(* Logix 5000 project; controller R400_500_XLS vendor 1 type 14 code 216 rev 31.11; software revision 31.01; part 2 of 32 *)

PROGRAM MainProgram   (* main routine MainRoutine *)
VAR
   Abort1 : DINT := 1;   // Not Used
        .0   // Initial step
        .1   // Remove stop condition
        .10   // Call module to fill sump Close Rcvry Tank Drain Valve
        .12   // Drain Rcvry Tank
        .14   // Call FC13 Drain Sump
        .16   // Sump draining phase is process
        .18   // Abort Completed Display Ready Mode screen
        .2   // No Recovery Tank Option or Recoverytank option and treament is Drying or Venting Reset Functions prior to drain sump
        .21   // Reset Functions
        .22   // Reset Functions prior to drain Rcvry Tank
        .24   // Reset Functions prior to drain sump
        .26   // Reset Functions prior to drain Rcvry Tank
        .28   // Reset Functions prior to drain sump
        .31   // Start Abort Sequence
        .4   // Check Filling Port
        .6   // Reset Functions prior to drain Rcvry Tank
        .8   // Reset Functions prior to fill sump
   Abort2 : SINT := 33;
        .0   // Initial Step
        .1   // Drying or Venting treatment is running Reset Functions prior to Vent Chamber
        .2   // Drying or Venting Treat. was running Exhaust Chamber (Abort Sequence) Enrg. Fan
        .5   // Initial Step
        .6   // Recirc. or F. Rinse Treat. was running Exhaust Chamber (Abort Sequence)
   Alarm : SINT := 1;   // Wait 3 seconds
        .0   // Initial step. No alarm detected.
        .1   // Alarm detected. Stop the cycle
        .2   // The alarm is acknowledged
        .3   // Display RESUME button
        .5   // Transition
        .6   // Transition
        .7   // Run mode
   AlarmAcked : BOOL;   // Alarm has been acked
   AlarmFlag : DINT;   // Active alarm flag
        .1   // Load door did not open flag
        .10   // Pure water tank safety water level reached
        .11   // Sump too long to fill
        .12   // Sump drain too long
        .13   // Sump too long to heat
        .14   // Sump RTD defective
        .15   // Sump temperature too high
        .16   // Pure water tank too long to fill
        .17   // Pure water tank drain too long
        .18   // Pure Water Tank too long to heat
        .19   // Pure Water Tank RTD defective
        .2   // Load door did not close flag
        .20   // Pure water tank temperature too high
        .21   // Pure water tank failed to dump
        .22   // Chemical Container 1 empty
        .23   // Chemical Container 2 empty
        .24   // Chemical Container 3 empty
        .25   // Chemical Container 4 empty
        .26   // Drying temperature not reached
        .27   // Chemical injection conductivity setpoint not reached
        .28   // Final rinse conductivity setpoint not reached
        .29   // Final rinse conductivity system defective
        .3   // Load door obstructed
        .30   // Chemcial conductivity system defective
        .31   // Pressure Transmitter defective
        .4   // Load door open
        .5   // Unload door did not open
        .6   // Unload door did not close
        .7   // Unload Door Obstructed
        .8   // Unload door Open
        .9   // Sump safety level reached
   AlarmFlag1 : DINT;
        .0   // Pump pressure too low
        .1   // Motor overload detected
        .10   // Waiting For Pure Water Filling Authorization
        .11   // Audit Trail Low Storage Memory
        .2   // Maintenance due
        .3   // Both doors open
        .4   // Drying RTD defective
        .5   // Master control relay deactivated
        .6   // PURE WATER TANK TEMPERATURE ABOVE TEMPERATURE RANGE ALLOWED
        .7   // PURE WATER TANK TEMPERATURE UNDER TEMPERATURE RANGE ALLOWED
        .8   // BATTERY LOW
        .9   // I/O Communication has been lost
   AlarmMuted : BOOL;
   AlarmTran0 : BOOL;   // Transition from step 3 to step 0
   Ashutdown : SINT := 1;   // Not Used
        .0   // Initial Step
        .1   // Call manual shutdown function Start signal from the automatic shutdown requirement
        .2   // Wait activation of Wake button (initial step of OPR-13)
        .3   // Enabled door printout and wait opening of the door
        .4   // Door is open
        .5   // Unloading completed
        .6   // Accept/Reject Cycle
   bAlrm : BOOL[64];
        [10]   // PURE WATER TANK TOO LONG TO DRAIN (trigger)
        [11]   // SUMP TOO LONG TO FILL (trigger)
        [12]   // SUMP TOO LONG TO HEAT (trigger)
        [13]   // SUMP DRAIN TOO LONG (trigger)
        [14]   // Chemical container 1 low
        [15]   // Chemical container 2 low
        [16]   // Chemical container 3 low
        [17]   // Chemical container 4 low
        [18]   // ALARM PURE WATER TANK TOO LONG TO FILL (trigger)
        [19]   // Pure water tank too long to heat
        [1]   // ALARM LOAD DOOR OBSTRUCTED (trigger)
        [20]   // ALARM PURE WATER TANK FAIL TO DUMP (trigger)
        [21]   // PURE WATER TANK TOO LONG TO DRAIN
        [22]   // Drying temperature not reached (trigger)
        [23]   // Chemical container 1 low
        [24]   // Chemical container 2 low
        [25]   // Chemical container 3 low
        [26]   // Chemical container 4 low
        [27]   // Conductivity is too long to reach set point
        [28]   // Final Rinse cond. sp not reached
        [29]   // Chemical container 1 low
        [2]   // ALARM LOAD DOOR DID NOT OPEN (trigger)
        [30]   // Chemical container 2 low
        [31]   // Chemical container 3 low
        [32]   // Chemical container 4 low
        [3]   // ALARM LOAD DOOR DID NOT CLOSE (trigger)
        [4]   // Reserved Load door open
        [5]   // ALARM UNLOAD DOOR OBSTRUCTED (trigger)
        [6]   // ALARM UNLOAD DOOR DID NOT OPEN (trigger)
        [7]   // ALARM UNLOAD DOOR DID NOT CLOSE (trigger)
        [8]   // Reserved Unload Door Open
        [9]   // SUMP TOO LONG TO DRAIN (trigger)
   bChangeFromNonHeatedToHeated : BOOL;
   bResetAllCycle : BOOL;
   bResetServiceMode : BOOL;
   CalCond : SINT;
        .1   // Calibration Enabled bit
        .2   // Wait for low calibration value
        .3   // Set Low value and Wait for High value
        .4   // Set High value and Verify Calibration
   CalFrinseCond : SINT;
        .1   // Calibration Enable bit
        .2   // Wait for low calibration value
        .3   // Set Low value and Wait for High value
        .4   // Set High value and Verify Calibration
   Calib : SINT;
        .0   // Enter Low Value
        .1   // Enter High Value
        .2   // Verify Calibration
   CalibCnt : SINT := 2;   // Calibration Step Counter
   CalibCondCnt : SINT;
   CalibData : UDT_SCALE[8] := ([0].InputMin := 213, [0].InputMax := 1207, [0].ScaledMin := 218.0, [0].ScaledMax := 1212.0, [0].DfInputMax := 1000, [0].DfScaledMax := 1000, [0].Input := 212, [0].Output := 21.7, [1].InputMin := 234, [1].InputMax := 1204, [1].ScaledMin := 239.0, [1].ScaledMax := 1210.0, [1].DfInputMax := 1000, [1].DfScaledMax := 1000, [1].Input := 222, [1].Output := 22.698767, [2].InputMin := 223, [2].InputMax := 1205, [2].ScaledMin := 228.0, [2].ScaledMax := 1210.0, [2].DfInputMax := 1000, [2].DfScaledMax := 1000, [2].Input := 214, [2].Output := 21.9, [3].InputMin := 4000, [3].InputMax := 20000, [3].ScaledMax := 60.0, [3].DfInputMin := 4000, [3].DfInputMax := 20000, [3].DfScaledMax := 60, [3].Input := 12566, [3].Output := 32.122498, [4].InputMin := 4000, [4].InputMax := 20000, [4].ScaledMax := 100.0, [4].DfInputMin := 4000, [4].DfInputMax := 20000, [4].DfScaledMax := 100, [4].Input := 9495, [4].Output := 34.34375, [5].InputMin := 4000, [5].InputMax := 20000, [5].ScaledMax := 100.0, [5].DfInputMin := 4000, [5].DfInputMax := 20000, [5].DfScaledMax := 100, [5].Input := 4000, [7].InputMin := 223, [7].InputMax := 1205, [7].ScaledMin := 228.0, [7].ScaledMax := 1210.0, [7].DfInputMax := 1000, [7].DfScaledMax := 1000, [7].Input := 302, [7].Output := 30.7);
        [0]   // Sump RTD Calibration data
        [1]   // Dry RTD Calibration data
        [2]   // PWT RTD Calibration data
        [3]   // Pressure Calibration data
        [4]   // Final Rinse Channel calibration data
        [5]   // Chemical Channe calibration data
        [6]   // Spare channel
        [7]   // Reserved for printouts
   CalibEnabled : BOOL;   // RTD Calibration Enabled bit
   CalibFrinseCondCnt : SINT;
   CalibIndex : DINT := 1;   // Calibration Pointer
   CalibPressCnt : SINT := 2;
   CalPressure : SINT;
   Change_PrintPtr_Value : BOOL;
   Chem_Pump : UDT_CHEM_PUMP[4] := ([0].FlowRate := 270, [1].FlowRate := 270, [2].FlowRate := 270, [3].FlowRate := 270);   // Chemical Pump flow rate
        [0].FlowRate   // Flow rate of Pump 1
        [1].FlowRate   // Flow rate of Pump 2
        [2].FlowRate   // Flow rate of Pump 3
        [3].FlowRate   // Flow rate of Pump 4
   CHEMICAL_COND_MAX_TIME : DINT := 360000;   // Timeout for the conductivity based chemical injection
   CHEMICAL_PUMP_OFF_TIME : DINT[4] := ([0] := 8, [1] := 8, [2] := 8, [3] := 8);
   CHEMICAL_PUMP_ON_TIME : DINT[4] := ([0] := 2, [1] := 2, [2] := 2, [3] := 2);
   ChemPumpIndex : DINT := 1;
   ChPumpRunningTime : REAL := 42.043003;
   ClearIndex : DINT := 300;
   Condenser : INT := 1025;
        .0   // Initial step. Condenser stopped
        .1   // Condenser operating
        .10   // Initial step. Condenser stopped
        .11   // Condenser operating
   CondenserHighFlow_1 : BOOL;   // Enables the condenser high flow valve
   CondenserHighFlow_2 : BOOL;   // Enables the condenser high flow valve
   CondenserLowFlow_1 : BOOL;   // Enables the condenser low flow valve
   CondenserLowFlow_2 : BOOL;   // Enables the condenser low flow valve
   CondenserTran : INT;
        .0   // From step 0 to 1
        .1   // From step 1 to 0
        .10   // From step 10 to step 11
        .11   // From step 11 to step 10
   Critical_Alarm : BOOL;
   CURRENT_CYCLE : DINT := 11;
   CustomCycleIterator : DINT := 11;
   CycExcBuffer : UDT_CYCLE := (PW[0].Wprt := 2, PW[0].Tmin := 1, PW[1].Wprt := 2, PW[2].Wprt := 2, PW[3].Wprt := 2, WSH[0].Wprt := 2, WSH[1].Wprt := 2, WSH[2].Wprt := 2, WSH[3].Wprt := 2, WSH[4].Wprt := 2, RINSE[0].Wprt := 2, RINSE[1].Wprt := 2, RINSE[2].Wprt := 2, RINSE[3].Wprt := 2, FRINSE.Tsec := 10, FRINSE.Drn := 1, DRY.HeatSensitive := 1, Lock := 1);
   CycleDryingStandard : UDT_DRY := (Mode := 1, Tmin := 15, HiLowTemp := 1);
   CycleModifBuffer : UDT_CYCLE := (PW[0].Wprt := 2, PW[0].Tmin := 1, PW[1].Wprt := 2, PW[2].Wprt := 2, PW[3].Wprt := 2, WSH[0].Wprt := 2, WSH[1].Wprt := 2, WSH[2].Wprt := 2, WSH[3].Wprt := 2, WSH[4].Wprt := 2, RINSE[0].Wprt := 2, RINSE[1].Wprt := 2, RINSE[2].Wprt := 2, RINSE[3].Wprt := 2, FRINSE.Tsec := 10, FRINSE.Drn := 1, DRY.HeatSensitive := 1, Lock := 1);
   CycleNotEmpty : SINT;
   Cycles : UDT_CYCLE[11] := ([0].PW[0].TrtNo := 1, [0].PW[0].Wprt := 1, [0].PW[0].Tmin := 2, [0].PW[1].Wprt := 2, [0].PW[2].Wprt := 2, [0].PW[3].Wprt := 2, [0].WSH[0].Wprt := 2, [0].WSH[0].Heat := 1, [0].WSH[0].Tmp := 65.6, [0].WSH[0].Tmin := 10, [0].WSH[0].ChemUsed_1 := 1, [0].WSH[0].ChemVol_1 := 4.0, [0].WSH[1].Wprt := 2, [0].WSH[2].Wprt := 2, [0].WSH[2].Heat := 1, [0].WSH[2].Tmp := 65.6, [0].WSH[2].Tmin := 1, [0].WSH[2].ChemUsed_1 := 2, [0].WSH[2].ChemVol_1 := 4.0, [0].WSH[3].Wprt := 2, [0].WSH[4].Wprt := 2, [0].RINSE[0].Wprt := 2, [0].RINSE[0].Tmin := 4, [0].RINSE[1].Wprt := 2, [0].RINSE[1].Tmin := 8, [0].RINSE[2].Wprt := 2, [0].RINSE[3].Wprt := 2, [0].FRINSE.Heat := 1, [0].FRINSE.Tmp := 50.0, [0].FRINSE.Tsec := 10, [0].FRINSE.Nb := 1, [0].FRINSE.Recirc := 1, [0].FRINSE.Drn := 1, [0].DRY.Mode := 1, [0].DRY.Tmin := 25, [0].DRY.HiLowTemp := 1, [0].Lock := 1, [1].PW[0].Wprt := 1, [1].PW[0].Tmin := 2, [1].PW[1].Wprt := 2, [1].PW[2].Wprt := 2, [1].PW[3].Wprt := 2, [1].WSH[0].Wprt := 2, [1].WSH[0].Heat := 1, [1].WSH[0].Tmp := 65.6, [1].WSH[0].Tmin := 10, [1].WSH[0].ChemUsed_1 := 1, [1].WSH[0].ChemVol_1 := 3.90625, [1].WSH[1].Wprt := 2, [1].WSH[2].Wprt := 2, [1].WSH[3].Wprt := 2, [1].WSH[4].Wprt := 2, [1].RINSE[0].Wprt := 2, [1].RINSE[0].Tmin := 4, [1].RINSE[1].Wprt := 2, [1].RINSE[1].Heat := 1, [1].RINSE[1].Tmp := 65.6, [1].RINSE[1].Tmin := 8, [1].RINSE[2].Wprt := 2, [1].RINSE[3].Wprt := 2,
        [1].FRINSE.Heat := 1, [1].FRINSE.Tmp := 65.6, [1].FRINSE.Tsec := 10, [1].FRINSE.Nb := 2, [1].FRINSE.Drn := 1, [1].DRY.HeatSensitive := 1, [1].Lock := 1, [2].PW[0].Wprt := 2, [2].PW[0].Tmin := 2, [2].PW[1].Wprt := 2, [2].PW[2].Wprt := 2, [2].PW[3].Wprt := 2, [2].WSH[0].Wprt := 2, [2].WSH[0].Heat := 1, [2].WSH[0].Tmp := 65.6, [2].WSH[0].Tmin := 10, [2].WSH[1].Wprt := 2, [2].WSH[2].Wprt := 2, [2].WSH[3].Wprt := 2, [2].WSH[4].Wprt := 2, [2].RINSE[0].Wprt := 2, [2].RINSE[0].Tmin := 4, [2].RINSE[1].Wprt := 1, [2].RINSE[1].Tmin := 8, [2].RINSE[2].Wprt := 2, [2].RINSE[3].Wprt := 2, [2].FRINSE.Tsec := 10, [2].FRINSE.Nb := 2, [2].FRINSE.Drn := 1, [2].DRY.Mode := 1, [2].Lock := 1, [3].PW[0].Wprt := 1, [3].PW[1].Wprt := 2, [3].PW[2].Wprt := 2, [3].PW[3].Wprt := 2, [3].WSH[0].Wprt := 2, [3].WSH[0].Heat := 1, [3].WSH[0].Tmp := 65.6, [3].WSH[0].ChemUsed_1 := 1, [3].WSH[0].ChemVol_1 := 0.9765625, [3].WSH[1].Wprt := 2, [3].WSH[2].Wprt := 2, [3].WSH[3].Wprt := 2, [3].WSH[4].Wprt := 2, [3].RINSE[0].Wprt := 2, [3].RINSE[1].Wprt := 2, [3].RINSE[2].Wprt := 2, [3].RINSE[3].Wprt := 2, [3].FRINSE.Heat := 1, [3].FRINSE.Tmp := 50.0, [3].FRINSE.Tsec := 30, [3].FRINSE.Recirc := 1, [3].FRINSE.Drn := 1, [3].DRY.Mode := 1, [3].DRY.Tmin := 25, [3].DRY.HiLowTemp := 1, [3].Lock := 1, [4].PW[0].Wprt := 2, [4].PW[0].Tmin := 2, [4].PW[0].Tsec := 30,
        [4].PW[1].Wprt := 1, [4].PW[1].Tmin := 1, [4].PW[2].Wprt := 2, [4].PW[3].Wprt := 2, [4].WSH[0].Wprt := 2, [4].WSH[0].Tmin := 10, [4].WSH[0].ChemUsed_1 := 1, [4].WSH[0].ChemVol_1 := 1.953125, [4].WSH[1].Wprt := 2, [4].WSH[1].Heat := 1, [4].WSH[1].Tmp := 65.6, [4].WSH[1].Tmin := 4, [4].WSH[2].Wprt := 2, [4].WSH[2].Tmin := 10, [4].WSH[2].ChemUsed_1 := 1, [4].WSH[2].ChemVol_1 := 3.90625, [4].WSH[3].Wprt := 2, [4].WSH[4].Wprt := 2, [4].RINSE[0].Wprt := 2, [4].RINSE[1].Wprt := 2, [4].RINSE[2].Wprt := 2, [4].RINSE[3].Wprt := 2, [4].FRINSE.Heat := 1, [4].FRINSE.Tmp := 50.0, [4].FRINSE.Tsec := 30, [4].FRINSE.Recirc := 1, [4].FRINSE.Drn := 1, [4].DRY.Mode := 1, [4].Lock := 1, [5].PW[0].Wprt := 2, [5].PW[1].Wprt := 2, [5].PW[2].Wprt := 2, [5].PW[3].Wprt := 2, [5].WSH[0].Wprt := 2, [5].WSH[0].Heat := 1, [5].WSH[0].Tmp := 65.6, [5].WSH[0].ChemUsed_1 := 2, [5].WSH[0].ChemVol_1 := 16.0, [5].WSH[1].Wprt := 2, [5].WSH[2].Wprt := 2, [5].WSH[3].Wprt := 2, [5].WSH[4].Wprt := 2, [5].RINSE[0].Wprt := 2, [5].RINSE[0].Tmin := 10, [5].RINSE[1].Wprt := 2, [5].RINSE[1].Tmin := 10, [5].RINSE[2].Wprt := 2, [5].RINSE[2].Tmin := 10, [5].RINSE[3].Wprt := 2, [5].FRINSE.Heat := 1, [5].FRINSE.Tmp := 50.0, [5].FRINSE.Tsec := 30, [5].FRINSE.Recirc := 1, [5].FRINSE.Drn := 1, [5].DRY.Mode := 1, [5].DRY.Tmin := 15, [5].DRY.HiLowTemp := 1, [5].Lock := 1, [6].PW[0].Wprt := 2, [6].PW[0].Tmin := 1,
        [6].PW[1].Wprt := 2, [6].PW[2].Wprt := 2, [6].PW[3].Wprt := 2, [6].WSH[0].Wprt := 2, [6].WSH[0].Heat := 1, [6].WSH[0].Tmp := 70.0, [6].WSH[0].ChemUsed_1 := 1, [6].WSH[0].ChemVol_1 := 1.953125, [6].WSH[1].Wprt := 2, [6].WSH[1].Tmin := 5, [6].WSH[1].ChemUsed_1 := 2, [6].WSH[1].ChemVol_1 := 1.953125, [6].WSH[2].Wprt := 2, [6].WSH[3].Wprt := 2, [6].WSH[4].Wprt := 2, [6].RINSE[0].Wprt := 2, [6].RINSE[1].Wprt := 2, [6].RINSE[2].Wprt := 2, [6].RINSE[3].Wprt := 2, [6].FRINSE.Tsec := 10, [6].FRINSE.MnNb := 1, [6].FRINSE.Drn := 1, [6].DRY.Mode := 1, [6].Lock := 1, [7].PW[0].Wprt := 2, [7].PW[0].Tmin := 1, [7].PW[1].Wprt := 2, [7].PW[2].Wprt := 2, [7].PW[3].Wprt := 2, [7].WSH[0].Wprt := 2, [7].WSH[1].Wprt := 2, [7].WSH[2].Wprt := 2, [7].WSH[3].Wprt := 2, [7].WSH[4].Wprt := 2, [7].RINSE[0].Wprt := 2, [7].RINSE[0].Heat := 1, [7].RINSE[0].Tmp := 80.0, [7].RINSE[0].Tmin := 1, [7].RINSE[1].Wprt := 2, [7].RINSE[2].Wprt := 2, [7].RINSE[3].Wprt := 2, [7].FRINSE.Heat := 1, [7].FRINSE.Tmp := 50.0, [7].FRINSE.Tsec := 10, [7].FRINSE.Nb := 1, [7].FRINSE.Drn := 1, [7].DRY.Mode := 1, [7].Lock := 1, [8].PW[0].Wprt := 2, [8].PW[0].Tmin := 1, [8].PW[1].Wprt := 2, [8].PW[2].Wprt := 2, [8].PW[3].Wprt := 2, [8].WSH[0].Wprt := 2, [8].WSH[1].Wprt := 2, [8].WSH[2].Wprt := 2, [8].WSH[3].Wprt := 2, [8].WSH[4].Wprt := 2, [8].RINSE[0].Wprt := 2, [8].RINSE[1].Wprt := 2,
        [8].RINSE[2].Wprt := 2, [8].RINSE[3].Wprt := 2, [8].FRINSE.Tsec := 10, [8].FRINSE.Drn := 1, [8].DRY.HeatSensitive := 1, [8].Lock := 1, [9].PW[0].Wprt := 2, [9].PW[1].Wprt := 2, [9].PW[2].Wprt := 2, [9].PW[3].Wprt := 2, [9].WSH[0].Wprt := 2, [9].WSH[1].Wprt := 2, [9].WSH[2].Wprt := 2, [9].WSH[3].Wprt := 2, [9].WSH[4].Wprt := 2, [9].RINSE[0].Wprt := 2, [9].RINSE[1].Wprt := 2, [9].RINSE[2].Wprt := 2, [9].RINSE[3].Wprt := 2, [9].FRINSE.Tsec := 10, [9].FRINSE.MnNb := 1, [9].FRINSE.Drn := 1, [9].DRY.Mode := 1, [9].Lock := 1, [10].PW[0].Wprt := 1, [10].PW[0].Tsec := 30, [10].PW[1].Wprt := 2, [10].PW[2].Wprt := 2, [10].PW[3].Wprt := 2, [10].WSH[0].Wprt := 2, [10].WSH[0].Tsec := 30, [10].WSH[0].ChemUsed_1 := 1, [10].WSH[0].ChemUsed_2 := 2, [10].WSH[0].ChemVol_1 := 1.0, [10].WSH[0].ChemVol_2 := 1.0, [10].WSH[1].Wprt := 2, [10].WSH[2].Wprt := 2, [10].WSH[3].Wprt := 2, [10].WSH[4].Wprt := 2, [10].RINSE[0].Wprt := 2, [10].RINSE[0].Heat := 1, [10].RINSE[0].Tmp := 65.5, [10].RINSE[0].Tsec := 30, [10].RINSE[1].Wprt := 2, [10].RINSE[2].Wprt := 2, [10].RINSE[3].Wprt := 2, [10].FRINSE.Heat := 1, [10].FRINSE.Tmp := 65.5, [10].FRINSE.Tsec := 10, [10].FRINSE.Nb := 1, [10].FRINSE.Drn := 1, [10].DRY.Mode := 1, [10].DRY.Tsec := 30, [10].DRY.HiLowTemp := 1, [10].Lock := 1);
        [0]   // EXTRA Care
   CyclesDefault : UDT_CYCLE[7] := ([0].PW[0].TrtNo := 1, [0].PW[0].Wprt := 2, [0].PW[0].Tmin := 1, [0].PW[1].Wprt := 2, [0].PW[2].Wprt := 2, [0].PW[3].Wprt := 2, [0].WSH[0].Wprt := 2, [0].WSH[0].Heat := 1, [0].WSH[0].Tmp := 65.6, [0].WSH[0].Tmin := 2, [0].WSH[0].Tsec := 30, [0].WSH[0].ChemUsed_1 := 1, [0].WSH[0].ChemVol_1 := 4.0, [0].WSH[1].Wprt := 2, [0].WSH[2].Wprt := 2, [0].WSH[2].Heat := 1, [0].WSH[2].Tmp := 65.6, [0].WSH[2].Tmin := 1, [0].WSH[2].ChemUsed_1 := 2, [0].WSH[2].ChemVol_1 := 4.0, [0].WSH[3].Wprt := 2, [0].WSH[4].Wprt := 2, [0].RINSE[0].Wprt := 2, [0].RINSE[0].Tsec := 30, [0].RINSE[1].Wprt := 2, [0].RINSE[1].Tsec := 30, [0].RINSE[2].Wprt := 2, [0].RINSE[3].Wprt := 2, [0].FRINSE.Heat := 1, [0].FRINSE.Tmp := 50.0, [0].FRINSE.Tsec := 30, [0].FRINSE.Nb := 1, [0].FRINSE.MnNb := 1, [0].FRINSE.Recirc := 1, [0].FRINSE.Drn := 1, [0].DRY.Mode := 1, [0].Lock := 1, [1].PW[0].Wprt := 2, [1].PW[1].Wprt := 2, [1].PW[2].Wprt := 2, [1].PW[3].Wprt := 2, [1].WSH[0].Wprt := 2, [1].WSH[0].Heat := 1, [1].WSH[0].Tmp := 54.0, [1].WSH[0].Tmin := 2, [1].WSH[0].ChemUsed_1 := 1, [1].WSH[0].ChemVol_1 := 2.0, [1].WSH[1].Wprt := 2, [1].WSH[2].Wprt := 2, [1].WSH[3].Wprt := 2, [1].WSH[4].Wprt := 2, [1].RINSE[0].Wprt := 2, [1].RINSE[0].Tsec := 15, [1].RINSE[1].Wprt := 2, [1].RINSE[2].Wprt := 2, [1].RINSE[3].Wprt := 2, [1].FRINSE.Heat := 1, [1].FRINSE.Tmp := 50.0, [1].FRINSE.Tsec := 30, [1].FRINSE.Nb := 1,
        [1].FRINSE.MnNb := 1, [1].FRINSE.Recirc := 1, [1].FRINSE.Drn := 1, [1].DRY.Mode := 1, [1].Lock := 1, [2].PW[0].Wprt := 2, [2].PW[0].Tmin := 2, [2].PW[1].Wprt := 2, [2].PW[2].Wprt := 2, [2].PW[3].Wprt := 2, [2].WSH[0].Wprt := 2, [2].WSH[0].Heat := 1, [2].WSH[0].Tmp := 54.0, [2].WSH[0].Tmin := 2, [2].WSH[0].ChemUsed_1 := 1, [2].WSH[0].ChemVol_1 := 4.0, [2].WSH[1].Wprt := 2, [2].WSH[2].Wprt := 2, [2].WSH[3].Wprt := 2, [2].WSH[4].Wprt := 2, [2].RINSE[0].Wprt := 2, [2].RINSE[0].Tsec := 30, [2].RINSE[1].Wprt := 2, [2].RINSE[2].Wprt := 2, [2].RINSE[3].Wprt := 2, [2].FRINSE.Heat := 1, [2].FRINSE.Tmp := 50.0, [2].FRINSE.Tsec := 30, [2].FRINSE.Nb := 1, [2].FRINSE.MnNb := 1, [2].FRINSE.Recirc := 1, [2].FRINSE.Drn := 1, [2].DRY.Mode := 1, [2].Lock := 1, [3].PW[0].Wprt := 1, [3].PW[0].Tmin := 2, [3].PW[1].Wprt := 2, [3].PW[2].Wprt := 2, [3].PW[3].Wprt := 2, [3].WSH[0].Wprt := 2, [3].WSH[0].Heat := 1, [3].WSH[0].Tmp := 65.6, [3].WSH[0].Tmin := 5, [3].WSH[0].ChemUsed_1 := 1, [3].WSH[0].ChemVol_1 := 4.0, [3].WSH[1].Wprt := 2, [3].WSH[2].Wprt := 2, [3].WSH[3].Wprt := 2, [3].WSH[4].Wprt := 2, [3].RINSE[0].Wprt := 2, [3].RINSE[0].Tmin := 1, [3].RINSE[1].Wprt := 2, [3].RINSE[1].Tmin := 1, [3].RINSE[2].Wprt := 2, [3].RINSE[3].Wprt := 2, [3].FRINSE.Heat := 1, [3].FRINSE.Tmp := 50.0, [3].FRINSE.Tsec := 10, [3].FRINSE.Nb := 1, [3].FRINSE.MnNb := 1,
        [3].FRINSE.Drn := 1, [3].DRY.Mode := 1, [3].DRY.Tmin := 15, [3].DRY.HiLowTemp := 1, [3].Lock := 1, [4].PW[0].Wprt := 2, [4].PW[1].Wprt := 2, [4].PW[2].Wprt := 2, [4].PW[3].Wprt := 2, [4].WSH[0].Wprt := 2, [4].WSH[1].Wprt := 2, [4].WSH[2].Wprt := 2, [4].WSH[3].Wprt := 2, [4].WSH[4].Wprt := 2, [4].RINSE[0].Wprt := 2, [4].RINSE[0].Tmin := 1, [4].RINSE[1].Wprt := 2, [4].RINSE[2].Wprt := 2, [4].RINSE[3].Wprt := 2, [4].FRINSE.Heat := 1, [4].FRINSE.Tmp := 50.0, [4].FRINSE.Tsec := 30, [4].FRINSE.Nb := 1, [4].FRINSE.MnNb := 1, [4].FRINSE.Recirc := 1, [4].FRINSE.Drn := 1, [4].DRY.Mode := 1, [4].Lock := 1, [5].PW[0].Wprt := 2, [5].PW[1].Wprt := 2, [5].PW[2].Wprt := 2, [5].PW[3].Wprt := 2, [5].WSH[0].Wprt := 2, [5].WSH[0].Heat := 1, [5].WSH[0].Tmp := 65.6, [5].WSH[0].Tmin := 10, [5].WSH[0].ChemUsed_1 := 2, [5].WSH[0].ChemVol_1 := 16.0, [5].WSH[1].Wprt := 2, [5].WSH[2].Wprt := 2, [5].WSH[3].Wprt := 2, [5].WSH[4].Wprt := 2, [5].RINSE[0].Wprt := 2, [5].RINSE[0].Tmin := 1, [5].RINSE[1].Wprt := 2, [5].RINSE[1].Tmin := 1, [5].RINSE[2].Wprt := 2, [5].RINSE[2].Tmin := 1, [5].RINSE[3].Wprt := 2, [5].FRINSE.Heat := 1, [5].FRINSE.Tmp := 50.0, [5].FRINSE.Tsec := 30, [5].FRINSE.Nb := 1, [5].FRINSE.MnNb := 1, [5].FRINSE.Recirc := 1, [5].FRINSE.Drn := 1, [5].DRY.Mode := 1, [5].Lock := 1, [6].PW[0].Wprt := 2, [6].PW[1].Wprt := 2,
        [6].PW[2].Wprt := 2, [6].PW[3].Wprt := 2, [6].WSH[0].Wprt := 2, [6].WSH[1].Wprt := 2, [6].WSH[2].Wprt := 2, [6].WSH[3].Wprt := 2, [6].WSH[4].Wprt := 2, [6].RINSE[0].Wprt := 2, [6].RINSE[1].Wprt := 2, [6].RINSE[2].Wprt := 2, [6].RINSE[3].Wprt := 2, [6].FRINSE.Tsec := 10, [6].FRINSE.MnNb := 1, [6].FRINSE.Drn := 1, [6].DRY.Mode := 1, [6].Lock := 1);   // Preliminary Data block to reset Cycles Values
        [0]   // EXTRACare
        [1]   // ENVIROCare
        [2]   // PLASTIC
        [3]   // STANDARD
        [4]   // RINSECare
        [5]   // DESCALER
        [6]   // CYCLE 7 to 11
   CycleSequence : UDT_CYCLE_SEQUENCE := (InitialStep := 1);
   CycleSmartDryingHeatSens : UDT_DRY := (HeatSensitive := 1);
   CycleSmartDryingRegular : UDT_DRY := (HiLowTemp := 1);
   CycleTime : DINT[11] := ([0] := 1489, [1] := 69, [2] := 1909, [3] := 2470, [4] := 1200, [5] := 120, [6] := 233, [7] := 960, [8] := 2027, [9] := 1140, [10] := 718);   // Last cycle time saved in seconds
   CycleUsageArraySize : DINT := 50;   // Size of the Cycle Usage Array
   CycleUsageDefaultUserName : STRING := '-';   // Default User Name
   CycleUsageDefaultValue : UDT_CYCLE_USAGE := (UserName := '-');
   CycleUsageFirstEmptyIndex : DINT := 50;   // Cycle Usage Array First Empty Index
   CycleUsageIterator : DINT;
   CycleUsagePrintoutCycleStartedCount : STRING := '2';
   CycleUsagePrintoutHeader : STRING := '*******  CYCLE USAGE  *******';
   CycleUsagePrintoutMessage : STRING := 'Cycle(s) Started';
   CycleUsagePrintoutSeparator : STRING := ' : ';
   CycleUsageSearchCurrentUser : BOOL;
   CycleUsageSearchFirstEmptyIndex : BOOL := 1;
   CycleWith_NonRecircFRinseDefault : UDT_FRINSE := (Heat := 1, Tmp := 50.0, Tsec := 10, Nb := 1, MnNb := 1, Drn := 1);
   CycleWith_RecircFRinseDefault : UDT_FRINSE := (Heat := 1, Tmp := 50.0, Tsec := 30, Nb := 1, MnNb := 1, Recirc := 1, Drn := 1);
   CycleWithoutDry : UDT_DRY := (Mode := 1);
   CycleWithoutFRinseWithoutTankDefault : UDT_FRINSE := (MnNb := 1, Recirc := 1, Drn := 1);
   CycleWithoutFRinseWithTankDefault : UDT_FRINSE := (Tsec := 10, MnNb := 1, Drn := 1);
   CycViewBuffer : UDT_WASH;
   Delta_T : REAL := 0.5;
   DESCALER : SINT := 5;
   DintBuffer : DINT[5] := ([0] := 3, [1] := 4);
   Drain_RcvryTnk_with_Sump : DINT := 1;   // 0 = Close Recovery Tank Drain Valve 1 = Open Recovery Tank Drain Valve
   DrainNo : DINT;
   DrnSmp : DINT := 1025;
        .0   // Initial Step
        .1   // CoolDown and Not Rcvry Tank option Low Water Volume
        .10   // Initial Step Recovery Tank is ready
        .11   // Performs Drain Type 3
        .12   // No Cooldown with Recovery Tank
        .13   // Perform Drain Type 3 Leave open Recovery Tank drain valve
        .14   // Perform Drain Type 3 Close Recovery Tank Drain Valve Water is saved in Recovery Tank
        .15   // Drain Recovery Tank
        .16   // Cooldown with Recovery Tank
        .17   // Performs Drain Type 1 or Drain Type 2 Leave open Recovery Tank drain valve
        .18   // Cooldown and not Recovery Tank Perform Drain Type 1 or Drain Type 2
        .19   // Perform Drain Type 3 Close Recovery Tank Drain Valve Water is saved in Recovery Tank
        .2   // CoolDown and Not Rcvry Tank option High Water Volume
        .20   // Start Rcvry Tank Cooldown seq. Fill Sump to cooldown Rcvry Tank
        .21   // Drain Recovery Tank and sump
        .28   // Rcvry Tank Cooldown seq. In progress
        .3   // Whitout cooldown Open Sump Drain Valve
        .4   // Start Sump Draining Timer
        .5   // Set Flag to exit module
        .6   // Retrun to step DrnSmp.0
        .7   // Open Cooldown valve
        .8   // Open Sump Drain Valve
        .9   // Open Condensate return Valve
   DRYING : DINT := 23;   // Drying id number
   DRYING_HEAT_SENSITIVE_SEL : DINT := 17;   // Drying heat sensitive
   DRYING_MODE_SEL : DINT := 14;   // Drying mode selector index
   drying_sp : REAL := 82.2;   // Drying temperature set point
   drying_sp_offset : REAL := 72.2;   // Low drying offset
   DRYING_TEMP_C_SEL : DINT := 15;   // Drying temperature index
   DRYING_TEMP_F_SEL : DINT := 16;   // Drying temperature index
   DRYING_TEMP_HIGH : REAL := 115.6;   // Smart drying high temperature set point
   DRYING_TEMP_LOW : REAL := 82.2;   // Smart drying low temperature set point
   DRYING_TEMP_STANDARD_LOW : REAL := 65.0;   // Regular drying low temperature set point
   DRYING_TIME_LONG : DINT := 20;   // Smart drying time for heat sensitive mode (in minute)
   DRYING_TIME_MIN_NUM : DINT := 11;   // Drying time (minutes) numeric input index
   DRYING_TIME_SEC_NUM : DINT := 12;   // Drying time (seconds) numeric input index
   DRYING_TIME_SHORT : DINT := 10;   // Smart drying time for heat regular mode (in minute)
   dryingSmartTime : DINT := 1200000;   // Duration of the smart drying phase
   DryingTempCool : REAL := 71.1;   // Temperature limit for the smart drying mode cooling phase
   DX_div_100 : REAL;
   ENVIRO_CARE : SINT := 1;
   EXTRA_CARE : SINT;
   F1rinse : DINT := 32769;   // Not Used
        .0   // Initial Step
        .1   // Print Treatment header
        .10   // Enable Final Rinse Evaluation
        .11   // Do another Final Rinse Returm to Frinse.1 step
        .12   // No more Final Rinse required Return to F1rinse.0 step
        .15   // Initial Step
        .16   // Fixed NB of Rinses Do Another Final Rinse Call Drain Sump
        .17   // Drain completed, Do another Final Rinse
        .18   // return to Step F1rinse.15
        .19   // Fixed NB of Rinses No more Final Rinse requested
        .20   // Drain Sump Last Final Rinse
        .21   // Set Water Saved flag
        .22   // No more final rinse required set flag to exit routine
        .23   // return to step F1rinse.15
        .3   // Call module to drain sump
        .5   // Fill Sump with Pure Water
        .7   // No Tank Recirc. PW Start Pump, heat sump recirc. timer
        .9   // Monitor Cond. Increment F. Rinse Cntr
   F2rinse : DINT := 1;   // Not Used
        .0   // Initial Step
        .1   // Print Final Rinse Header
        .11   // End of Heating Start Water Transfer
        .13   // Tank, N-R Final Rinse Start Pump (Low Speed)
        .15   // Add 1 to Nb of Final Rinse Done
        .16   // Fixed NB of Rinses Do Another Final Rinse Call Drain Sump
        .17   // Enable Final Rinse Evaluation
        .18   // Do another Final Rinse return to F2rinse.1
        .19   // No More Final Rinse is required. return to step F2rinse.0
        .20   // Initial Step
        .21   // Cycle is stopped Wait Resume
        .23   // Trig Alarm Pure Water Tank Failed To Dump
        .3   // Call Module to drain sump
        .5   // Call to fill Pure Water Tank
        .7   // Check if treatment is heated
        .9   // Call Module to Heat Pure Water Tank
   F3rinse : DINT := 1;   // Not Used
        .0   // Initial Step
        .1   // Print Final Rinse Header
        .11   // End of Heating Gravity Transfer Step
        .13   // Delay to close valve
        .15   // Tank Recirc. Final Rinse Start Pump, Heat Sump, Enable Recirc. Timer
        .17   // Add 1 to Number of Final Rinse Done
        .18   // Enable Grafcet Evaluation
        .19   // Another Final Rinse is required. return to step F3rinse.1
        .20   // No More Final Rinse is required. return to step F3rinse.0
        .21   // Trig Alarm Pure Water Tank Failed To Dump
        .3   // Call module to drain sump
        .5   // Call module to fill pure water tank
        .7   // Check if treatment is heated
        .9   // Call module to Heat Pure Water Tank
   F4rinse : INT := 1;   // Transition for the conductivity based evalutaion
        .0   // Initial step.
        .1   // Save the water conductivity.
        .10   // Another rinse is required
        .2   // Drain the sump. Close the transfer valve.
        .3   // Another rinse is required
        .4   // Check Final Rinse Drain setting
        .5   // Drain the sump.
        .6   // Sump does not need to be drained.
        .7   // No more final rinse required
        .8   // Set the alarm.
        .9   // Drain the sump.
   F4rinse_Tran : INT;   // Transitions for the conductivity based evaluation
        .0   // Step 0 => Step 1
        .1   // Step 1 => Step 2
        .10   // Step 1 => Step 8
        .11   // Step 8 => Step 9
        .12   // Step 9 => Step 10
        .13   // Step 10 => Step 0
        .2   // Step 2 => Step 3
        .3   // Step 3 => Step 0
        .4   // Step 1 => Step 4
        .5   // Step 4 => Step 5
        .6   // Step 5 => Step 7
        .7   // Step 4 => Step 6
        .8   // Step 6 => Step 7
        .9   // Step 7 => Step 0
   FC05_ONS : DINT;
   FC06_ONS : DINT;
   FC06Tran1 : BOOL;   // Condition for the wash treatment to start
   FC07Tran1 : BOOL;   // Condition for the rinse treatment to start
   FC22_SumpWaterVolume : REAL := 47.3;   // Water volume
   FC22_Tran1 : BOOL;   // First transition
   FC22_Tran3 : BOOL;   // Third transition
   FC22_Tran4 : BOOL;   // Fourth transition
   FC22_WashIndex : SINT := 2;
   FC23_BaseConductivity : REAL := 1.4172212;   // Base conductivity of the water prior to the injection
   FC23_ChemicalPumpIndex : DINT := 2;   // Chemical pump index
   FC23_CompensatedSetPoint : REAL;   // Injection compensated chemical conductivity
   FC23_FinalConductivity : REAL := 13.218668;   // Final value of the chemical conductivity
   FC23_OffsetSetPoint : REAL;   // Set point before enabling the on/off sequence
   FC23_ONS : SINT := 2;
   FC23_StartSignal : BOOL;   // Conductivity based chemical injection
   FC23_WashIndex : DINT := 2;   // Current index of the wash treatment
   FC45_NextMaintDate : DINT[3] := ([0] := 2090, [1] := 8, [2] := 14);   // Next maintenance due date
        [0]   // Next maintenance due -Year-
        [1]   // Next maintenance due -Month-
        [2]   // Next maintenance due -Day-
   FC65_Enabled_signal : BOOL;   // Enables the treatment evaluation
   FC65_Treatment_counter : DINT;   // Treatment counter
   FC83_AutoSpeed : BOOL;   // Cycle pump speed selection
   FC83_AutoWtrLevel : BOOL;   // Cycle water level selection
   FC83_CyclePerm : BOOL := 1;   // Cycle permission selection
   FC83_DryHeatSensitive : DINT := 1;   // Drying is heat sensitive?
   FC83_DryTemp : DINT;   // Drying temperature (hi/low)
   FC83_FRinse_Drained : DINT := 1;   // Drained final rinse flag
   FC83_FRinse_Heated : DINT;   // Heated final rinse flag
   FC83_FRinse_Recirculated : DINT;   // Recirculated final rinse flag
   FC83_ONS : SINT := -106;
   FC87_CalibChemPmp : SINT;   // Calibration chemical pumps activation bits
        .0   // Chemical pump 1 toggle bit
        .1   // Activate chemical pump 1 output
        .2   // Chemical pump 2 toggle bit
        .3   // Activate chemical pump 2 output
        .4   // Chemical pump 3 toggle bit
        .5   // Activate chemical pump 3 output
        .6   // Chemical pump 4 toggle bit
        .7   // Activate chemical pump 4 output
   FC87_CalibChemPmpMsg : SINT := 1;   // Chemical pump calibration step message
        .0   // Press start button to begin the injection
        .1   // Injection in progress...
        .2   // Enter chemical volume injected
   FC87_ChemCalibRemainTime : DINT := 40;
   FC87_ChemPumpIndex : SINT;   // Index of the selected chemical pump to calibrate
   FC87_LastValue : SINT;
   FC87_ONS : DINT;
   Fill_Sump : DINT := 32769;
        .0   // Initial Step
        .1   // Set Alarm time Enrg. Cold Water Valve
        .10   // PW Filling Request
        .11   // PW Draining Deadleg
        .15   // Initial Step (Heating)
        .16   // Enrg Sump Steam Valve (SumpTemp < 26.6 C)
        .17   // Pre-Heating Enrg Sump Steam Valve (SumpTemp < 37.7 C)
        .18   // Stop Heating
        .19   // Return to step Fill_Smp.15
        .2   // Set Alarm Time Enrg. Hot Water Valve
        .3   // Set Alarm time Enrg. Pure Water valve
        .4   // Sump is full Wait Step
        .5   // Set Flag to exit module
        .6   // Flag is reset
        .7   // Set Alarm Time Enrg. Hot Water Valve
        .8   // Set Alarm Time Enrg. Hot Water Valve
   FINAL_RINSE_MAX_NBR : INT := 9;   // Maximum nimber of final rinse
   FINALRINSE_1 : DINT := 14;   // Final rinse 1 id number
   FINALRINSE_2 : DINT := 15;   // Final rinse 2 id number
   FINALRINSE_3 : DINT := 16;   // Final rinse 3 id number
   FINALRINSE_4 : DINT := 17;   // Final rinse 4 id number
   FINALRINSE_5 : DINT := 18;   // Final rinse 5 id number
   FINALRINSE_6 : DINT := 19;   // Final rinse 6 id number
   FINALRINSE_7 : DINT := 20;   // Final rinse 7 id number
   FINALRINSE_8 : DINT := 21;   // Final rinse 8 id number
   FINALRINSE_9 : DINT := 22;   // Final rinse 9 id number
   First_Inj_conc : BOOL;
   First_PwWshRnseTtr : DINT := 1;
   FRINSE_COND_SET_POINT_NUM : DINT := 18;   // Final rinse conductivity set point numeric input index
   FRINSE_DRAIN_SEL : DINT := 19;   // Final rinse drained selector's index
   FRINSE_HEATING_SEL : DINT := 18;   // Final rinse heating selector's index
   FRINSE_MIN_NUMBER_NUM : DINT := 17;   // Final rinse minimum number of final rinse numeric input index
   FRINSE_NUMBER_NUM : DINT := 16;   // Final rinse number of final rinse numeric input index
   FRINSE_RECIRC_SEL : DINT := 20;   // Final rinse recirculated selector's index
   FRINSE_TIME_MIN_NUM : DINT := 14;   // Final rinse time (minutes) numeric input index
   FRINSE_TIME_SEC_NUM : DINT := 15;   // Final rinse time (seconds) numeric input index
   FRINSE_TYPE_SEL : DINT := 21;   // Final rinse type selector's index
   FRinseCondValue : REAL := 1.0062485;   // Stored value of the conductivity
   H0_Temp : REAL := 64.0;
   H1_Temp : REAL := 64.0;
   HDelta_T : REAL := 6.0999985;
   HeatSmp : DINT := 1049601;
        .0   // Initial Step
        .1   // Enrg Sump steam valve (continuously)
        .10   // Initial Step
        .11   // Enrg. Sump Heating contactor (continuous)
        .12   // Stop Heating
        .13   // Enrg. Sump Heating contactor for xx sec
        .2   // Enrg Sump steam valve 2 sec.
        .20   // Initial step
        .21   // Set Recir. Hys.Value
        .22   // Start recirculation Timer
        .23   // Stop Recirculation Timer
        .24   // Recirculation Time is elapsed
        .25   // Re-initialize HeatSmp.20 step
        .26   // Non Heated PW-W-R With Hot Water Port and Heat Recovery Tank option
        .27   // Stop Pre-Heating
        .28   // Pre-heating Energized Sump Steam Valve
        .3   // De-enrg Sump steam valve 4 sec.
        .4   // Wait termperature change
        .5   // Enrg. Sump Steam Valve or Electric Contactor
   HighLimt : REAL := 0.1;
   I_0_Missing : BOOL;
   I_Pw_Tnk_Lvl_Sw_Deb : BOOL;   // Debounced pure water tank level switch (100ms)
   iBuffer : DINT[5] := ([1] := 30, [4] := 9);
   iDecimalSeparatorIndex : INT := 5;
   iFindCRLFIndex : INT := 21;   // Index Of CRLF in String
   iIndexClearMessageOverflowBuffer : INT := 300;   // Message Overflow Buffer is sPrntArray(200-300)
   Inj_Cond : SINT := 1;   // Conductivity injection based steps
        .0   // Initial step
        .1   // Wait for temperature.
        .2   // Compute the set point.
        .3   // Conductivity based chemical injection. Start the pump.
        .4   // Conductivity based chemical injection. On/off routine.
        .5   // End of injection.
   Inj_Cond_Tran : SINT;   // Conductivity injection based transitions
        .0   // Step 0 => 1
        .1   // Step 1 => 2
        .2   // Step 2 => 3
        .3   // Step 3 => 4
        .4   // Step 4 => 5
        .5   // Step 5 => 0
   Inj_Time : SINT := 1;   // Time based chemical injection steps
        .0   // Initial step
        .1   // Computes the injection time required;starts the chemical pump;starts the timer.
        .2   // Resets the injection timer
        .3   // Computes the injection time required;starts the chemical pump;starts the timer.
        .4   // Resets the injection timer
   InjMan : SINT := 1;
        .0   // Manual injection has not started yet
        .1   // Manual injection in progress
   L310ER_Led : DINT := 3;
   Last_Hdelta_T : REAL := 6.0999985;
   Last_PwWshRnseTtr : DINT := 11;
   LowLimt : REAL;
   LowPressAlmSp : REAL := 5.0;   // Pump pressure too low setpoint
   M : DINT[5] := ([0] := 2304, [1] := 4100, [3] := 4, [4] := 1024);   // Memory Bits
        [0].0   // Door Safety (Futur E-Stop if required)
        [0].1   // Cmd_Opn_Ld_Dr
        [0].10   // Cycle in process bit
        [0].11   // Door(s) are closed
        [0].12   // Start Treatment evaluation
        [0].13   // Start treatment
        [0].14   // End of Pre-Wash Treatment
        [0].15   // Initiate Module (Abort)
        [0].16   // Initiate Module (Abort)
        [0].17   // End of sump filling sequence (FC11)
        [0].18   // Shelf is not present
        [0].19   // Shelf is present
        [0].2   // Cmd_Clse_LdDr
        [0].20   // Pulse start pump low speed
        [0].21   // Enrg. pump Low Speed Service Mode
        [0].22   // Pulse start pump high Speed Service Mode
        [0].23   // Enrg. pump High Speed Service Mode
        [0].24   // Service Mode Pump Low Speed
        [0].25   // Service Mode Pump High Speed
        [0].26   // Start Sump Heating (Pulse)
        [0].27   // Reset Grafcet (Abort, enf of recirc.)
        [0].28   // Flag End of Recirc. phase
        [0].29   // Service Mode Enabled
        [0].3   // Cmd_Opn_Unld_Dr
        [0].30   // Start Sump draining phase
        [0].31   // Initiate after Abort
        [0].4   // Cmd_Cls_Unld_Dr
        [0].5   // 1= Open Sump Drain Valve
        [0].6   // 1 = Final Rinse Treatment present in cycle
        [0].7   // 1= Open Pure Water Outlet Valve
        [0].8   // Sump is drained
        [0].9   // Initiate Module (Abort)
        [1].0   // Flag End of Sump Draining phase
        [1].1   // Rcvry Tank Module (End of sump draining phase)
        [1].10   // Interlock Bit
        [1].11   // End of Final Rinse Fixed Number of Rinses
        [1].12   // Drying Treatment in cycle
        [1].13   // Interlock Bit
        [1].14   // start 1st N-R Final Rinse Treatment
        [1].15   // Cycle is started (1st treatment is a final rinse)
        [1].16   // Initiate module WSH_57 (Abort)
        [1].17   // End of rinse treatment flag
        [1].18   // Manual injection is over
        [1].19   // End of venting flag
        [1].2   // Supervisor mode enabled
        [1].20   // Initiate Module (Abort)
        [1].21   // End of drying
        [1].22   // Enrg drying heater
        [1].23   // Drying temperature set point reached in smart drying mode
        [1].24   // Drying Treatment Enrg drying fan
        [1].25   // Enrg drying isolation valve
        [1].26   // Drying Enrg transfer valve
        [1].27   // Enrg. Pure water tank Fill valve
        [1].28   // Start filling the pure water tank
        [1].29   // The pure water tank is full (signal for FC08 Module)
        [1].3   // End of wash phase
        [1].30   // A cycle has started and a final rinse is programmed and the thank is full
        [1].31   // Activate the steam valve
        [1].4   // Start Recvry Tank Cooling Phase
        [1].5   // Initiate module (Abort)
        [1].6   // Initiate Module (Abort)
        [1].7   // End of time based chemical injeciton
        [1].8   // Initiate Module (Abort)
        [1].9   // start 1st Final Rinse Treatment
        [2].0   // Activate the electric element
        [2].1   // The pure water tank has reached the set point
        [2].10   // Set PLC and HMI Date and time flag
        [2].11   // Start calibration chemical pump
        [2].12   // Chemical pump calibration in progress
        [2].13   // End chemical pump calibration
        [2].14   // Battery Low Interlock
        [2].16   // Shutdown Unit Water in Recovery Tank, Drain Rcvry Tank and Sump
        [2].17   // Shutdown Unit No Water in Recovery Tank, Drain Sump
        [2].18   // Init. Grafcet First scan or Test cancelled
        [2].2   // Initiate Module (Abort)
        [2].3   // Maintenance due flag
        [2].4   // Maintenance Due Interlock
        [2].5   // Detects the falling edge of the sump heating signal
        [2].6   // Initialize sequence
        [2].7   // End of conductivity injection
        [2].8   // End of conductivity based final rinse
        [2].9   // Set HMI Date and Time flag
        [3].0   // Interlock Bit
        [3].1   // Start 1st R. Final Rinse with PWT
        [3].10   // Sump Temp. too High Open sump drain valve 1 min
        [3].11   // PWT Temp. too High Open sump drain valve and PWT outlet valve for 1 min
        [3].12   // Sump Heating rate low
        [3].13   // Enable Visiblity of numeric pad
        [3].14   // WSH_30 Print Treatment Pump Pressure
        [3].15   // Set initial value
        [3].16   // WSH-41 Print footer
        [3].17   // WSH-22, Drain sump Enrg Dry Fan and Iso valve
        [3].18   // Door maintenance WSH-64 Disable Unload Door Open Alarm
        [3].19   // Initiate Module (Abort)
        [3].2   // Functions are reset
        [3].20   // Audible alarm request
        [3].21   // Enrg audible alarm continuously
        [3].22   // From SPV-18 Enrg. audible alarm output
        [3].23   // Automatic Shutdown enabled
        [3].24   // Print Calib Data
        [3].25   // Print Hardware option
        [3].26   // Print System option
        [3].27   // Enrg. Audible alarm
        [3].28   // Enrg. Audible alarm
        [3].29   // Enrg Close then Open pilot valve at next activation
        [3].3   // Abort in Process
        [3].30   // Energ. Close then Open Coil
        [3].31   // Close door at next button activation
        [3].4   // Iniate end of neutralization printout
        [3].5   // Init Alarm.0
        [3].6   // 1= Close Heat Recovery Tank Drain Valve
        [3].7   // Thermal Schock Risk Pure Water Tank Temp > SumpTemp
        [3].8   // Thermal Schock Risk SumpTemp > Pure Water Tank Temp
        [3].9   // 1st treatment is a final rinse treatment
        [4].0   // Enrg. Close pilot valve
        [4].10   // Initial Step
        [4].11   // Service Mode Enrg Hot Water Fill valve
        [4].12   // Service Mode Enrg Hot Water Fill valve
        [4].13   // Service Mode Enrg Hot Water fill valve
        [4].2   // Enrg Close then Open pilot valve at next activation
        [4].3   // Energ. Close then Open Coil
        [4].4   // From screen 18 Ready Mode
        [4].5   // From screen 30 Analog input
   MaxPressRecord : REAL;
   MaxTrtTempSp : REAL := 95.03;
   MinorFaultCheck : TIMER := (PRE := 30000, ACC := 17512, EN := 1, TT := 1);
   MinorFaultRecord : FaultRecord;
   MinPressRecord : REAL;
   NbFinalRinseDone : DINT;
   Neutral : SINT := 1;
        .0   // Initial Step
        .1   // Inject Neutralizant
        .2   // Start Recirc.pump
        .3   // End of neutralization
        .4   // Start delay to stop pump
        .5   // Inject Neutralizant
        .7   // Keep Pump Running
   NeutralizantPump : SINT;
   NeutralizationInjTime : DINT := 23949;
   NeutralizationPhaseRequired : BOOL;
   NeutralizationRecircTime : DINT;
   New_Value : SINT;
   NON_RECIRCULATED_FINAL_RINSE_MINUTES : DINT;   // Number of minutes for the non recirculated final rinse
   NON_RECIRCULATED_FINAL_RINSE_SECONDS : DINT := 10;   // Number of seconds for the non recirculated final rinse
   OneShot : DINT[1] := ([0] := 8389760);
   ONS_FC01 : DINT := 8;
   ONS_FC05 : DINT;
   ONS_FC07 : SINT;
   ONS_FC08 : DINT := 2048;
   ONS_FC09 : SINT;
   ONS_FC11 : DINT;
   ONS_FC12 : DINT := 256;
   ONS_FC13 : DINT := 64;
   ONS_FC17_1 : BOOL;
   ONS_FC17_2 : BOOL;
   ONS_FC22 : SINT;
   ONS_FC24 : SINT := 2;
   ONS_FC25 : DINT;
   ONS_FC34 : DINT;
   ONS_FC37 : DINT;
   ONS_FC39 : DINT;
   ONS_FC40 : SINT;
   ONS_FC45 : DINT;
   ONS_FC64 : DINT;
   ONS_FC65 : DINT;
   ONS_FC84 : SINT;
   ONS_FC85 : SINT := 16;
   ONS_FC86 : DINT := 292;
   ONS_SPV17 : SINT := 16;
   ONS_WSH30 : SINT := 4;
   ONS_WSH35 : SINT := 1;
   OPR_16_TreatPrint_Ptr : DINT;
   PLASTIC_CARE : SINT := 2;
   PresetMin : SINT;
   PresetSec : SINT := 30;
   PREWASH_1 : DINT := 1;   // Pre-wash 1 id number
   PREWASH_2 : DINT := 2;   // Pre-wash 2 id number
   PREWASH_3 : DINT := 3;   // Pre-wash 3 id number
   PREWASH_4 : DINT := 4;   // Pre-wash 4 id number
   PreWash_Select : BOOL;
   PrewashIndex : SINT := 1;   // Index of the selected pre-wash treatment
   PreWtrDrnTme : DINT := 10000;
   PrimeChemPmp : SINT;   // Prime chemical pumps activation bits
        .0   // Chemical pump 1 toggle bit
        .1   // Activate chemical pump 1 output
        .2   // Chemical pump 2 toggle bit
        .3   // Activate chemical pump 2 output
        .4   // Chemical pump 3 toggle bit
        .5   // Activate chemical pump 3 output
        .6   // Chemical pump 4 toggle bit
        .7   // Activate chemical pump 4 output
   Print_Data : BOOL;   // Print Treatment data
   print_Door_opened_template : STRING := 'DOOR OPENED:';   // Template for the door opened message
   print_Footer_template : STRING[7] := ([0] := 'CYCLE COMPLETED:', [1] := 'TOTAL CYCLE TIME:', [2] := 'READY TO UNLOAD...', [3] := 'MINIMUM PRESSURE:', [4] := 'MAXIMUM PRESSURE:', [5] := 'PSIG', [6] := 'Bar');   // Template for the cycle footer
   print_Header_template : STRING[6] := ([0] := 'CYCLE NAME:', [1] := 'DATE:', [2] := 'START TIME:', [3] := 'CYCLE COUNTER:', [4] := 'SERIAL NUMBER:', [5] := 'USER:');   // Template for the cycle header
   Print_Speed_Water : BOOL;
   Print_TreatEnd_Start_Data : BOOL;   // 2nd treatment of the cycle is started, pirnt Treatment Completed and Treatment data
   Print_TreatStart_Data : BOOL;   // Cycle is started Print start time and treatment data of the first treatment of the cycle
   PrintBufferInjectionRate : REAL;
   PrintCalibdata : STRING[9] := ([0] := '**********  CALIBRATION DATA  **********', [1] := 'UNIT SERIAL NUMBER:', [2] := 'LOW RAW:', [3] := 'HIGH RAW:', [4] := 'LOW VALUE:', [5] := 'HIGH VALUE:', [6] := '***  CHEMICAL PUMPS FLOW RATE  ***', [7] := 'mL/min', [8] := ': ');
   printCycleParameters : STRING[2] := ([0] := 'CYCLE PARAMETERS', [1] := 'CYCLE:');
   printNeutralization : STRING[5] := ([0] := 'NEUTRALIZATION COMPLETED');
   PrintoutMSGTranslation : DINT := 1;   // Grapcet for Printout Message Translation
        .0   // Initial step of messages transfer
        .1   // Start a message transfer
        .2   // Send a message transfer request
        .3   // Message received
        .4   // Message transfer completed
   PrintoutMSGTranslationONS : INT;
   PrintPressureDelay : DINT := 5000;
   PrintSensorName : STRING[7] := ([0] := '***  SUMP RTD  ***', [1] := '***  DRY RTD  ***', [2] := '***  PWT RTD  ***', [3] := '***  PRESSURE CHANNEL  ***', [4] := '***  F. R. CHANNEL  ***', [5] := '***  CHEMICAL CHANNEL  ***');
   printTreatString : STRING[85] := ([0] := 'FINAL RINSE 1', [1] := 'PRE-WASH 1', [2] := 'PRE-WASH 2', [3] := 'PRE-WASH 3', [4] := 'PRE-WASH 4', [5] := 'WASH 1', [6] := 'WASH 2', [7] := 'WASH 3', [8] := 'WASH 4', [9] := 'WASH 5', [10] := 'RINSE 1', [11] := 'RINSE 2', [12] := 'RINSE 3', [13] := 'RINSE 4', [14] := 'FINAL RINSE 1', [15] := 'FINAL RINSE 2', [16] := 'FINAL RINSE 3', [17] := 'FINAL RINSE 4', [18] := 'FINAL RINSE 5', [19] := 'FINAL RINSE 6', [20] := 'FINAL RINSE 7', [21] := 'FINAL RINSE 8', [22] := 'FINAL RINSE 9', [23] := 'DRYING', [28] := 'TEMPERATURE:', [29] := 'REGULAR', [30] := 'TREATMENT START:', [31] := 'WATER PORT:', [32] := 'HOT WATER', [33] := 'COLD WATER', [34] := 'PURE WATER', [35] := 'TREAT. TEMP:', [36] := 'NON-HEATED', [37] := 'DEG$B0C', [38] := 'DEG$B0F', [39] := 'TREATMENT TIME:', [40] := 'CHEMICAL USED:', [41] := 'NONE', [46] := 'MANUAL', [47] := 'INJECTION TYPE:', [48] := 'TIME BASED', [49] := 'TREATMENT COMPLETED:', [50] := 'CONDUCTIVITY', [51] := 'CONCENTRATION:', [52] := 'oz/gal', [53] := 'ml/L', [54] := '0.0', [55] := 'CONDUCTIVITY SETPOINT:', [56] := 'mS/cm', [57] := 'LAST RINSE DRAIN:', [58] := 'YES', [59] := 'NO', [60] := 'RECIRCULATED:', [61] := 'FINAL RINSE TYPE:', [62] := 'FIXED NUMBER', [63] := 'CONDUCTIVITY', [64] := 'NUMBER OF FINAL RINSE:', [65] := 'MIN. NUMBER OF FINAL RINSE:', [66] := 'CONDUCTIVITY SETPOINT:', [67] := ' $B5S/cm',
        [68] := 'MODE:', [69] := 'SMART', [70] := 'STANDARD', [71] := 'TEMPERATURE: LOW (65.0 DEG$B0C)', [72] := 'TEMPERATURE: HIGH (115.6 DEG$B0C)', [73] := 'TEMPERATURE: LOW (149.0 DEG$B0F)', [74] := 'TEMPERATURE: HIGH (240.0 DEG$B0F)', [75] := 'HEAT SENSITIVE', [76] := 'FINAL RINSE', [77] := 'PUMP SPEED:', [78] := 'AUTO', [79] := 'LOW', [80] := 'WATER LEVEL:', [81] := 'HIGH', [82] := 'F. RINSE COND. VALUE:', [83] := 'CHEMICAL COND. VALUE:', [84] := 'PUMP PRESSURE :');   // Treatment String
        [0]   // Buffer
        [42]   // Not Used
        [43]   // Not Used
        [44]   // Not Used
        [45]   // Not Used
        [54]   // Concentration Value pinrt buffer
        [67]   // micro character Hexa value
   PumpLowFRinse : DINT := 3000;   // Delay for pump low speed during final rinse treatment
   PumpLowPW_W_R : DINT := 5000;   // Delay for pump low speed during pre-wash, wash and rinse treatments
   PURE_WATER_HEATING_TIME : DINT := 1200000;   // Time before an alarm is thrown when the pure water tank is heating
   PureWaterTankFilling : BOOL;   // Start PWT filling
   PW_HeatSp_5 : REAL := -5.0;
   PW_HeatSp_X : REAL := 5.0;
   PwExcBuffer : UDT_PW := (TrtNo := 1, Wprt := 2, Tmin := 1);
   PWHeat : SINT := 1;
        .1   // Energ. Sump Steam Valve (Continuous)
        .2   // Start Off delay
        .3   // Energ Steam Valve 2 sec.
        .4   // Temp Change too High steam valve is not activated
        .5   // Setpoint is reached
   PWR_PrintBuffer : UDT_WASH := (Wprt := 2, Tsec := 30, InjType_2 := 1);
   PWR_UP : DINT := 256;
        .0   // Initial Step Displayed screen 7
        .1   // Allow to close doors
        .2   // Door(s|) are pressurized
        .3   // Start Power-up drain
        .4   // Drain Sump
        .5   // Water detected in Sump
        .6   // Drain Pure Water Tank
        .7   // Water Detected in Pure Water Tank
        .8   // Power-Up Completed
   PWTnkTempAlmSp : REAL := 98.03;   // Pure water tank temperature too high setpoint
   rBuffer : REAL[4] := ([0] := 50.0, [1] := 50.051, [2] := 1.0, [3] := 50.0);
   Rcvry_Tnk_Tmp : REAL;   // Water Temperature of the Heat Recovery Tank
   RecircLowHysteresis : REAL := 49.0;
   ResetCycleName : BOOL;
   ResetMute : BOOL;
   rIn_WSH61 : REAL := 50.0;
   RINSE_1 : DINT := 10;   // Rinse 1 id number
   RINSE_2 : DINT := 11;   // Rinse 2 id number
   RINSE_3 : DINT := 12;   // Rinse 3 id number
   RINSE_4 : DINT := 13;   // Rinse 4 id number
   RINSE_CARE : SINT := 4;
   Rinse_Select : BOOL;
   RinseExcBuffer : UDT_RINSE := (Wprt := 2, Tsec := 30);
   RinseIndex : SINT := 1;
   RLO : BOOL;   // Logic result
   Run : DINT := 4100;
        .1   // Cycle is Started
        .10   // Ready to Unload No auto shutdown
        .11   // Door is open
        .12   // WSH-58 Unloading completed
        .13   // Accept/Reject Cycle
        .2   // Run/Stop bit 1 = Cycle is not paused 0 = Cycle is paused
        .3   // Stop Cycle
        .4   // Remove Stop Condtion
   s00_Nb : STRING := '00';
   s0_Nb : STRING := '0';
   s2lastdigits : STRING := '01';
   s36 : STRING := '36';
   s360 : STRING := '360';
   s3600 : STRING := '3600';
   s36000 : STRING := '36000';
   s360000 : STRING := '360000';
   s3600000 : STRING := '3600000';
   s36000000 : STRING := '36000000';
   s360000000 : STRING := '360000000';
   sCRLF : STRING := '$0D$0A';
   sDecimalSeparator : STRING := '.';
   sDigits1_2 : STRING := '60';
   Second_Inj_conc : BOOL;
   sEmptyString : STRING;   // Used on HMI(DO NOT DELETE)
   Service : DINT[2] := ([0] := 256);   // Unused Service Mode Memory Bit
        [0]   // Used Service Mode Memory Bit
        [0].0   // Used Service Mode Memory Bit
        [0].1   // Used Service Mode Memory Bit
        [0].10   // Used Service Mode Memory Bit
        [0].11   // Stop Door Operation
        [0].12   // Used Service Mode Memory Bit
        [0].13   // Used Service Mode Memory Bit
        [0].14   // Used Service Mode Memory Bit
        [0].15   // Used Service Mode Memory Bit
        [0].16   // Used Service Mode Memory Bit
        [0].17   // Used Service Mode Memory Bit
        [0].18   // Used Service Mode Memory Bit
        [0].19   // Used Service Mode Memory Bit
        [0].2   // Used Service Mode Memory Bit
        [0].20   // Used Service Mode Memory Bit Start HW filling
        [0].21   // Used Service Mode Memory Bit
        [0].22   // Used Service Mode Memory Bit
        [0].23   // Used Service Mode Memory Bit
        [0].24   // Used Service Mode Memory Bit
        [0].25   // Used Service Mode Memory Bit
        [0].26   // Used Service Mode Memory Bit
        [0].27   // Used Service Mode Memory Bit
        [0].28   // Used Service Mode Memory Bit
        [0].29   // Used Service Mode Memory Bit
        [0].3   // Used Service Mode Memory Bit
        [0].30   // Used Service Mode Memory Bit
        [0].31   // Used Service Mode Memory Bit
        [0].4   // Used Service Mode Memory Bit
        [0].5   // Used Service Mode Memory Bit
        [0].6   // Used Service Mode Memory Bit
        [0].7   // Used Service Mode Memory Bit
        [0].8   // free
        [0].9   // Stop Door Operation
        [1]   // Unused Service Mode Memory Bit
        [1].0   // Used Service Mode Memory Bit
        [1].1   // Used Service Mode Memory Bit
        [1].10   // Used Service Mode Memory Bit
        [1].11   // Used Service Mode Memory Bit
        [1].12   // Used Service Mode Memory Bit
        [1].13   // Used Service Mode Memory Bit
        [1].14   // Used Service Mode Memory Bit
        [1].15   // Used Service Mode Memory Bit
        [1].16   // Used Service Mode Memory Bit
        [1].17   // Used Service Mode Memory Bit
        [1].18   // Used Service Mode Memory Bit
        [1].19   // Used Service Mode Memory Bit
        [1].2   // Used Service Mode Memory Bit
        [1].20   // Used Service Mode Memory Bit
        [1].21   // Used Service Mode Memory Bit
        [1].22   // Used Service Mode Memory Bit
        [1].23   // Used Service Mode Memory Bit
        [1].3   // Used Service Mode Memory Bit
        [1].4   // Used Service Mode Memory Bit
        [1].5   // Used Service Mode Memory Bit
        [1].6   // Used Service Mode Memory Bit
        [1].7   // Used Service Mode Memory Bit
        [1].8   // Used Service Mode Memory Bit
        [1].9   // Used Service Mode Memory Bit
   ServicePassword : DINT := 160;   // Service Password
   SET_POINT_FRACTION : REAL[4] := ([0] := 0.8, [1] := 0.8, [2] := 0.8, [3] := 0.8);
   sFll_Zero : STRING[20] := ([0] := '0');
   Shutdown : SINT := 1;   // Shutdown sequence steps
        .0   // Initial step
        .1   // Drain the sump and the recovery tank.
        .2   // Drain the pure water tank.
        .3   // The shutdown sequence is over
   Shutdown_Tran : SINT;   // Shutdown sequence transitions
        .0   // Step 0 => Step 1
        .1   // Step 1 => Step 2
        .2   // Step 2 => Step 3
        .3   // Step 1 => Step 3
        .4   // Step 3 => Step 0
   sInvertedPairs : STRING := '0160';
   sLastdigit : STRING := '14526001';
   SMART_MODE_DRYING_HEATCOOL_SEC : DINT := 900;   // Heating and cooling time constant for the smart mode drying (sec.)
   sMessageToPrint : STRING := 'DOOR OPENED:14:17:14$0D$0A';   // Message To Print
   SmpDrnTme : DINT := 10000;
   SmpHeatingSp : REAL := 50.0;
   SmpLowHysteresis : REAL := 48.0;
   sOut_WSH61 : STRING := '50.0';
   sPrntArray : STRING[300];   // Printer String Array
   SRE3_Serial_Number : STRING := '3614526001';   // Serial number
   sResetPrinter : STRING := '$00$1B#P$00$1B@';   // Clears Printer buffer jplv04f ASCII
   Srl_Prt : SERIAL_PORT_CONTROL := (LEN := 19, POS := 19, EU := 1, DN := 1, EM := 1);   // Serial Port Control
   sSpaceCharacter : STRING := ' ';   // Space Character
   STANDARD : SINT := 3;
   start_1 : SINT := 5;
   start_2 : SINT := 7;
   StartPump1 : BOOL;   // Pump Low Speed
   StartPump2 : BOOL;   // Pump High Speed
   StartPump3 : BOOL;   // Main Pump running
   sTempo1 : STRING := '22.0';
   sTempo2 : STRING := '14526001';
   String : STRING[50] := ([0] := '-', [1] := '2026', [2] := '08', [3] := '17', [4] := '17-', [5] := '17-08', [6] := '17-08-', [7] := 'Mail Sent Successfully.', [8] := '11', [9] := ' ', [10] := '02', [11] := ' ', [12] := '10', [13] := ' ', [14] := ':', [15] := '11:', [16] := '11:02', [17] := '11:02:', [18] := ' ', [19] := '  -  ', [20] := '17-08-2026  -  ', [21] := '50.0509987', [22] := '.', [23] := ' ', [24] := 'MAINTENANCE DUE', [25] := 'DOOR OPENED:14:17:14$0D$0A$0D$0A');   // String
        [0]   // _ Dash Characters
        [10]   // Min String
        [11]   // Email ActiveX Failure Code
        [12]   // Sec String
        [13]   // Email Command String
        [14]   // : colon string
        [15]   // string buffer
        [16]   // string buffer
        [17]   // string buffer
        [18]   // Cell Phone + Domain
        [19]   // string buffer
        [1]   // Year string
        [20]   // string buffer
        [22]   // Period char.
        [23]   // To Email Address
        [24]   // DataStore Plus String Input
        [25]   // Printer String Output
        [2]   // Month String
        [3]   // Day String
        [4]   // string buffer
        [5]   // string buffer
        [6]   // string buffer
        [7]   // Mail Sent Successfully
        [8]   // Hour String
        [9]   // Blank Space String
   String_Temp : STRING := '1';
   SUMP_HIGH_VOLUME_400 : REAL := 36.0;   // High sump volume
   SUMP_HIGH_VOLUME_500 : REAL := 47.3;
   SUMP_LOW_VOLUME_400 : REAL := 22.0;   // Low sump volume
   SUMP_LOW_VOLUME_500 : REAL := 28.4;
   SumpHeatingStopped : BOOL;   // Sump heating falling edge
   SumpTempAlmSp : REAL := 98.03;   // Sump temperature too high setpoint
   SumpWaterVolume : DINT := 1;   // Sump Water Volume 0 =Low 1= High
   Supervisor : DINT;
        .0   // Supervisor memory bit
   T0_Temp : REAL := 49.9;
   T1_Temp : REAL := 49.9;
   TempChange : BOOL;
   tHandshakeToggle : TIMER := (PRE := 6000);
   Tmr : TIMER[107] := ([0].PRE := 2000, [1].PRE := 3000, [2].PRE := 20000, [3].PRE := 120000, [4].PRE := 90000, [4].ACC := 90000, [4].EN := 1, [4].DN := 1, [5].PRE := 10000, [6].PRE := 10000, [7].PRE := 120000, [8].PRE := 100, [9].PRE := 1000, [10].PRE := 40000, [11].PRE := 5000, [12].PRE := 3000, [13].PRE := 100, [14].PRE := 100, [15].PRE := 2000, [16].PRE := 4000, [17].PRE := 5000, [18].PRE := 1800000, [19].PRE := 100, [20].PRE := 30000, [21].PRE := 75000, [22].PRE := 2000, [23].PRE := 10000, [24].PRE := 2100, [25].PRE := 45000, [26].PRE := 45000, [27].PRE := 42044, [28].PRE := 3000, [29].PRE := 10000, [30].PRE := 15000, [31].PRE := 120000, [32].PRE := 30000, [33].PRE := 30000, [34].PRE := 5000, [35].PRE := 1200000, [36].PRE := 120000, [37].PRE := 480000, [38].PRE := 100, [39].PRE := 4000, [40].PRE := 1200000, [41].PRE := 3000, [42].PRE := 2500, [43].PRE := 45000, [44].PRE := 60000, [45].PRE := 120000, [46].PRE := 1200000, [47].PRE := 2000, [48].PRE := 60000, [49].PRE := 2000, [50].PRE := 8000, [51].PRE := 5000, [52].PRE := 360000, [53].PRE := 1000, [54].PRE := 3000, [55].PRE := 1000, [56].PRE := 10000,
        [57].PRE := 500, [58].PRE := 500, [59].PRE := 2000, [59].ACC := 2000, [60].PRE := 100, [61].PRE := 1000, [62].PRE := 100, [63].PRE := 100, [64].PRE := 10000, [65].PRE := 60000, [66].PRE := 1200000, [67].PRE := 40000, [69].PRE := 1000, [70].PRE := 60000, [71].PRE := 2000, [72].PRE := 1000, [73].PRE := 15000, [74].PRE := 5000, [75].PRE := 2000, [76].PRE := 3000, [77].PRE := 1000, [78].PRE := 3000, [80].PRE := 1000, [81].PRE := 1000, [82].PRE := 2000, [83].PRE := 2000, [84].PRE := 2000, [85].PRE := 2000, [86].PRE := 2000, [87].PRE := 60000, [88].PRE := 20000, [89].PRE := 6000, [90].PRE := 2000, [91].PRE := 7000, [92].PRE := 3000, [93].PRE := 2000000, [94].PRE := 23949, [95].PRE := 15000, [97].PRE := 1250, [99].PRE := 5000, [100].PRE := 2000, [101].PRE := 3000, [102].PRE := 2000, [103].PRE := 500, [104].PRE := 500, [105].PRE := 100, [106].PRE := 100);
        [0]   // Email Alarms Timer
        [100]   // Debounce delay
        [101]   // Delay between printouts
        [102]   // Delay Mag Door
        [103]   // Delay to switch from close to open coil
        [104]   // Delay to switch from close to open coil
        [105]   // Debouncing Delay (same delay as automatic mode)
        [106]   // Debouncing Delay (same delay as automatic mode)
        [10]   // Heating Timer (Filling sump)
        [11]   // Delay to switch to high speed
        [12]   // Delay to switch from low to high speed
        [13]   // Delay to de-energize
        [14]   // Delay to de-energize
        [15]   // Delay steam valve on
        [16]   // Delay steam valve off
        [17]   // Enrg Sump Heating contactor for xx sec
        [18]   // Sump Heating Alarm Timer
        [1]   // Email Timer
        [20]   // Recirculation Timer
        [21]   // Sump Draining Timer
        [22]   // Delay for lost of door sensor signal
        [23]   // Audible alarm delay
        [24]   // On-Off Timer Pilot Light Alternate Green and Red connection
        [25]   // Rcvry Tank/Sump Draining Timer
        [26]   // Rcvry Tank Drain Timer #1
        [27]   // Time Based Injection Timer
        [28]   // Delay to Open Pure Water Tank Outlet valve
        [29]   // Non-Recirclation Delay
        [2]   // Email Timeout
        [30]   // Trnasfer Water Gravity Delay
        [31]   // Vapor removal timer
        [32]   // Drying Timer (Time/Temperature modue)
        [33]   // Drying fan delay
        [34]   // Drying timer delay
        [35]   // Drying element timer
        [36]   // Drying cooling delay (Time/Temperature mode)
        [37]   // Pure water tank filling alarm
        [38]   // Debounce timer
        [39]   // Off delay Timer
        [3]   // Email Command Timeout
        [40]   // Alarm timer (bAlrm[19])
        [41]   // Alarm sequence delay to let the HMI see the trigger = 0
        [42]   // Closing Valve delay
        [43]   // Delay to drain the Rcvry Tank
        [44]   // Venting Delay
        [45]   // Recirc. or F. Rinse Treat. was running Exhaust Chamber (Abort Sequence)
        [46]   // Condenser timer
        [46].ACC   // Condenser counter variable
        [47]   // Condenser timer
        [48]   // Pure water tank drain timer
        [49]   // Conductivity injection on time
        [4]   // Power-up Dealy
        [50]   // Conductivity injection off time
        [51]   // Debouncing delay Conductivity set point reached
        [52]   // Conductivity based Alarm timer
        [53]   // Cycle time second counter
        [57]   // Interlock delay with Pure Water Tank Steam valve
        [58]   // Interlock delay with Sump Steam Valve
        [59]   // Delay after which, valve closes
        [5]   // Delay to Drain Sump
        [61]   // Cycle time wizard one second timer
        [62]   // Sump temperature too high timer
        [63]   // Pure water tank temperature too high timer
        [64]   // Pump pressure too low timer
        [65]   // Open valves on high temperature alarm timer
        [67]   // Chemical pump calibration timer
        [68]   // Sump Level Switch Debouncing delay
        [69]   // PWT Level Switch Debouncing delay
        [6]   // Delay to Drain Pure Water Tank
        [70]   // Comm alarm delay
        [71]   // 2 sec. delay to enrg. steam valve
        [72]   // Delay to print alarm
        [73]   // Delay for Water Stabilization
        [7]   // Sump Fill Alarm Timer
        [87]   // Sump heating rate delay
        [88]   // Heating interval alarm timer
        [89]   // Delay to display new password value before closing numeric pad entry
        [8]   // Debounce Sump Low Level Switch
        [90]   // Delay for pressure stabilization
        [91]   // Delay for mixing water
        [92]   // Timer Door Safety Test End
        [94]   // Neutralizant Injection Timer
        [95]   // Recirc. Timer
        [97]   // JPLV06
        [99]   // Delay to stop pump
        [9]   // String Copy Debounce
   Treatment_info : DINT;   // Treatment message conditions
        .4   // Heating message conditions
   TreatmentPrint_Ptr : SINT;
   TrecircSec : DINT := 30;
   Trt_Drying : SINT := 1;
        .0   // Initial step
        .1   // Drain the sump
        .2   // Open/close the valves
        .3   // Standard Mode drying routine
        .4   // Standard Mode Time based cooling
        .5   // Smart drying routine
        .6   // Smart Drying Temperature based cooling
        .7   // End of the drying phase
   Trt_Drying_Tran : INT;
        .0   // Step 0 => step 1
        .1   // Step 0 => step 2
        .2   // Step 1 => step 2
        .3   // Step 2 => step 3
        .4   // Step 3 => step 4
        .5   // Step 4 => step 7
        .6   // Step 2 => step 5
        .7   // Step 5 => step 6
        .8   // Step 6 => step 7
        .9   // Step 0 => step 7
   Trt_PrWsh : DINT := 1;
        .0   // Initial Step
        .1   // Call Fill Sump
        .2   // Start Pump, heat Enable drain of Recovery Tank
        .3   // Wait Step
        .4   // Call Drain Sump
        .5   // Sump draining and Recovery Tank draining phase completed
        .6   // Return to initial step
   Trt_Rinse : DINT := 1;   // Rinse steps
        .0   // Initial step
        .1   // Fill the sump
        .2   // Start pump, start heating, start recirculation
        .3   // Wait the recovery tank
        .4   // Starts the draining phase
        .5   // Rinse treatement over
        .6   // One scan delay
   Trt_Vapor_Exhaust : BOOL;   // Vapor exhaust fan is on
   Trt_Wsh : DINT := 1;
        .0   // Initial Step
        .1   // Sump Filling, Injection time based
        .2   // Filling done
        .3   // Manual chemical injection (FC24)
        .4   // Sump Heating, Start Pump
        .5   // Conductivity based injection, Start recirculation timer
        .6   // Check if neutralization is required
        .7   // Start sump draining
        .8   // End of wash treatment
   Unld_Door : DINT;
        .0   // Initialization
        .10   // Initial Step Open/Close Unload Door
        .11   // Enrg. Unload Door Open Pilot Valve
        .12   // Door is open Keep enrg. Unload Door Open Pilot Valve
        .13   // Trig Alarm Unlad Door Did Not Open
        .14   // Enrg. Unoad Door Close Pilot Valve
        .15   // Door is closed Keep enrg. Unload Door close Pilot Valve
        .16   // Trig Alarm Unload Door Did Not Close
        .17   // Trig Alarm Unload Door Obstructed
   USER_DEFINED_10 : SINT := 9;
   USER_DEFINED_11 : SINT := 10;
   USER_DEFINED_7 : SINT := 6;
   USER_DEFINED_8 : SINT := 7;
   USER_DEFINED_9 : SINT := 8;
   VENTING : DINT := 24;   // Venting id number
   VolumeInjected_ML : REAL := 189.19351;
   VolumeNeutralizer : REAL := 189.19351;
   WASH_1 : DINT := 5;   // Wash 1 id number
   WASH_2 : DINT := 6;   // Wash 2 id number
   WASH_3 : DINT := 7;   // Wash 3 id number
   WASH_4 : DINT := 8;   // Wash 4 id number
   WASH_5 : DINT := 9;   // Wash 5 id number
   Wash_Select : BOOL;
   washerMode : SINT := 1;   // Washer Mode Flag 0 -> Ready; 1 -> Supervisor; 2 -> Service; 3 -> Run.
   WashIndex : SINT;
   WashInjectionType1 : DINT;
   WaterSaved : BOOL;   // Water Saved In Sump (Last Final Rinse Water)
   WSH36_CycleTimePercentage : DINT := 100;
   WSH36_SecondsRemaining : DINT;
   WSH36_TotalMinutesRemaining : DINT;
   WSH36_TotalSecondsRemaining : DINT;
   WSH41_Door_opened : STRING := 'DOOR OPENED:14:17:14$0D$0A';
   WSH41_End_signal : BOOL;   // End of cycle signal
   WSH41_Header : STRING[6] := ([0] := 'CYCLE NAME:EXTRACare', [1] := 'DATE:14-08-2026', [2] := 'START TIME:13:52:02', [3] := 'CYCLE COUNTER:60', [4] := 'SERIAL NUMBER:3614526001', [5] := 'USER:service');   // The header being transferred to the print queue.
   WSH41_Hour : DINT;
   WSH41_Minute : DINT := 24;
   WSH41_ONS : SINT;
   WSH41_Second : DINT := 49;
   WSH41_Start_signal : BOOL;   // Start cycle signal One shot rising edge
   WSH41_Temp_time : STRING[3] := ([0] := '00', [1] := '24', [2] := '49');
   WSH41_Time_template : STRING := ':';
   WSH41_Total_minute : DINT;
   WSH41_Total_second : DINT;
   WSH41_Total_time : STRING := '00:24:49';
   WSH41_Zero : STRING := '0';
   WSH56_StartHeating : BOOL;   // Start heating
   WSH56_StartPump : BOOL;   // Start pump signal
   WSH56_StartRecirculation : BOOL;   // Start the recirculation
   WSH56_TreatmentInfo : BOOL;   // Treatment information for the conductivity injection
   WSH61_Footer : STRING[6] := ([0] := 'CYCLE COMPLETED:14:16:52', [1] := 'TOTAL CYCLE TIME:00:24:49', [2] := 'READY TO UNLOAD...');   // The footer being transferred to the print queue.
   WSH_35 : BOOL;   // End of neutralization phase
   WshExcBuffer : UDT_WASH := (Wprt := 2, Heat := 1, Tmp := 65.6, Tmin := 1, ChemUsed_1 := 2, ChemVol_1 := 4.0);
   Zero_Value : SINT := 1;
END_VAR
